FUNCTION_BLOCK FB_CoverState IMPLEMENTS I_CoverState
VAR_INPUT
END_VAR
VAR_OUTPUT
END_VAR
VAR
	pCover : POINTER TO FB_CoverControl;
END_VAR

{warning 'add method implementation '}
METHOD CloseCommand : BOOL
END_METHOD

METHOD FB_init : BOOL
VAR_INPUT
	bInitRetains : BOOL; // if TRUE, the retain variables are initialized (warm start / cold start)
	bInCopyCode : BOOL;  // if TRUE, the instance afterwards gets moved into the copy code (online change)
	pCover : POINTER TO FB_CoverControl;
END_VAR
THIS^.pCover := pCover;
END_METHOD

{warning 'add method implementation '}
METHOD OpenCommand : BOOL
END_METHOD

{warning 'add method implementation '}
METHOD RunState : BOOL
END_METHOD

{warning 'add method implementation '}
METHOD StopCommand : BOOL
END_METHOD

{warning 'add method implementation '}
METHOD SuccessfulFinished : BOOL
END_METHOD

END_FUNCTION_BLOCK

(* stored: Version 1.1.0.1, ProductVersion 3.1.4024.15
   POU FB_CoverState: Id {ca7d5149-bdab-48ed-9905-85ea4e750734}, SpecialFunc None
   Method CloseCommand: Id {195a36c7-9415-4524-9a5c-92ace990b07a}
   Method FB_init: Id {23c9b3ea-154f-4df6-949c-573bcf58c403}
   Method OpenCommand: Id {93a49747-2f23-4c26-96ad-cf4c3a310ea8}
   Method RunState: Id {a75daf41-ae92-4270-96c0-c0e432dac00e}
   Method StopCommand: Id {74a48edf-d297-4f18-80dd-9a1ebdef05c5}
   Method SuccessfulFinished: Id {4605a4e0-f930-436f-87ef-999f307c9f93} *)
